                  Waypoint OP_PowderA_abov: TCP in base x=-12.145 y=-363.335 z=315.326 mm, rx=-0.7771 ry=1.753 rz=-1.7409 rad; joints [-58.232, -116.012, -83.989, -160.83, 75.01, 1.147] deg; TCP offset x=0 y=0 z=161 mm, rx=3.1415 ry=0 rz=0 rad
                  Waypoint OP_PowderA_pick: TCP in base x=-12.145 y=-363.335 z=179.899 mm, rx=-0.7771 ry=1.753 rz=-1.7409 rad; joints [-58.242, -124.732, -92.401, -143.702, 75.051, 1.161] deg
                  URCap Gripper (Robotiq_Grippers, Robotiq Inc.) dataModel(position=100.0, force=30.19607843137255, speed=30.19607843137255, positionInDouble=100.0, forceInDouble=30.19607843137255, speedInDouble=30.19607843137255, slaveIds=[9], blocking=true)
                  Wait Sleep waitTime=0.5
                  Set DigitalOutput pin=GRP_3F_Open; digitalValue=1
                  SuppressedNode
                    Script: Motors_off()
                  Waypoint OP_PowderA_abov: motionParameters(jointSpeed=1.047198 jointAcceleration=1.396263 cartesianSpeed=0.05 cartesianAcceleration=0.3); TCP in base x=-12.145 y=-363.335 z=315.326 mm, rx=-0.7771 ry=1.753 rz=-1.7409 rad; joints [-58.232, -116.012, -83.989, -160.83, 75.01, 1.147] deg
                  Waypoint Op_PowA_wP: TCP in base x=-173.728 y=-372.934 z=295.117 mm, rx=-0.9724 ry=1.541 rz=-1.5487 rad; joints [-67.269, -106.894, -99.849, -153.52, 49.211, 1.028] deg
              URCap Approach Pose (SensoPart VISOR Robotic, SensoPart Industriesensorik GmbH) dataModel(visorOffsetZ=0.0, visorJointSpeed=25.0, visorJointAcc=30.0); state(isChildrenLocked=true)
              URCap Target Pose (SensoPart VISOR Robotic, SensoPart Industriesensorik GmbH) dataModel(visorToolSpeed=50.0, visorToolAcc=100.0); state(isChildrenLocked=true)
              Folder Close Gripper
                target_pose := pose_add(get_actual_tcp_pose(), p[0,0,-0.1,0,0,0])
                MoveL speed 250 mm/s, acceleration 1200 mm/s^2 (useActiveTCP=true optimoveEnabled=false optiMoveSpeed=0.3 optiMoveAcceleration=0.09) feature=Base
                  Waypoint Variable (Variable): motionParameters(jointSpeed=1.047198 jointAcceleration=1.396263 cartesianSpeed=0.05 cartesianAcceleration=0.3); variable(name=target_pose)
                URCap Gripper (Robotiq_Grippers, Robotiq Inc.) dataModel(position=0.0, force=30.19607843137255, speed=30.19607843137255, positionInDouble=0.0, forceInDouble=30.19607843137255, speedInDouble=30.19607843137255, slaveIds=[9], blocking=true)
              URCap Exit Pose (SensoPart VISOR Robotic, SensoPart Industriesensorik GmbH) dataModel(visorOffsetZ=0.0); state(isChildrenLocked=true)
            URCap No Object Detected (SensoPart VISOR Robotic, SensoPart Industriesensorik GmbH) dataModel(Variable(key=visorNoObjCountVar, variable(name=easyPickNoObj_7, initializeExpression=0)))
              Popup Message (haltProgram=false message=No weigh scale detected inputType=Text)
        place_pose := get_actual_tcp_pose()
        Script: center_pose()
        SuppressedNode
          center_tilt_pos := P_center
        MoveJ speed 60 deg/s, acceleration 80 deg/s^2 (useActiveTCP=true optimoveEnabled=false optiMoveSpeed=0.3 optiMoveAcceleration=0.09) feature=Base
          Waypoint Waypoint_1: TCP in base x=-451.049 y=-340.589 z=308.224 mm, rx=0.0971 ry=0.091 rz=-1.5784 rad; joints [-127.334, -100.578, -80.109, -94.907, 86.186, -126.663] deg
    Case (caseValue=42)
      Folder Powder Emptying
        Script: zero_scale()
        Task := "Emptying"
        SuppressedNode
          URCap VISOR Robotic App (SensoPart VISOR Robotic, SensoPart Industriesensorik GmbH) dataModel(visorAppTemplate=1); state(isChildrenLocked=true)
            URCap Easy Pick Setup (SensoPart VISOR Robotic, SensoPart Industriesensorik GmbH) dataModel(visorId=0, visorSetJob=true, visorImageAcqSetup=2, visorCalibSetNo=9, visorDetector=1, visorOffsetSet=true, visorImageAcqSource=2, visorJobName=Weigh_target, visorSetupStatus=5, Pose(key=visorGripPose, Position(key=posePosition, Length(key=X value=-0.477246 unit=M), Length(key=Y value=0.05319 unit=M), Length(key=Z value=0.184004 unit=M)), Rotation(key=poseRotation, Angle(key=RX value=0.786642 unit=RAD), Angle(key=RY value=1.426517 unit=RAD), Angle(key=RZ value=-0.850311 unit=RAD))), Feature(key=visorImageAcqFeature name=FRM_Centrifuge)); state(isChildrenLocked=true)
            URCap Process (SensoPart VISOR Robotic, SensoPart Industriesensorik GmbH) dataModel(Variable(key=visorCounterVar, variable(name=easyPickCount_4, initializeExpression=0)), Variable(key=visorPartsFoundVar, variable(name=easyPickParts_4, initializeExpression=0))); state(isChildrenLocked=true)
              URCap Image Acquisition Pose (SensoPart VISOR Robotic, SensoPart Industriesensorik GmbH) state(isChildrenLocked=true)
              URCap Object Detected (SensoPart VISOR Robotic, SensoPart Industriesensorik GmbH) state(isChildrenLocked=true)
                Folder Open Gripper
                  Script: tare_scale()
                  Wait Sleep waitTime=0.2
                  Weight_value := get_weight()
                  Wait Sleep waitTime=0.2
                  Script: compute_level_percent(W_now, Weight_value)
                  If level≥10.0
                    MoveJ speed 60 deg/s, acceleration 80 deg/s^2 (useActiveTCP=true optimoveEnabled=false optiMoveSpeed=0.3 optiMoveAcceleration=0.09) feature=Base
                      Waypoint Spatula_otw: TCP in base x=-38.472 y=-263.141 z=425.351 mm, rx=-0.0004 ry=-0.0001 rz=3.0344 rad; joints [-68.119, -57.773, -97.702, -114.504, 90.127, 27.957] deg
                      Waypoint pick_spat_L_abv: TCP in base x=247.376 y=-151.301 z=298.406 mm, rx=0 ry=-0.0005 rz=3.0677 rad; joints [-4.058, -56.828, -117.366, -95.794, 90.156, 90.183] deg
                    MoveL speed 250 mm/s, acceleration 1200 mm/s^2 (useActiveTCP=true optimoveEnabled=false optiMoveSpeed=0.3 optiMoveAcceleration=0.09) feature=Base
                      Waypoint spat_L_pick: TCP in base x=244.425 y=-151.048 z=192.288 mm, rx=0 ry=-0.0005 rz=3.0677 rad; joints [-4.109, -56.947, -132.87, -80.171, 90.162, 90.196] deg
                      URCap Gripper (Robotiq_Grippers, Robotiq Inc.) dataModel(position=100.0, force=30.0, speed=0.0, positionInDouble=100.0, forceInDouble=30.0, speedInDouble=0.0, slaveIds=[9], blocking=true)
                      Waypoint spat_L_lift: TCP in base x=247.5 y=-151.291 z=242.147 mm, rx=0 ry=-0.0005 rz=3.0677 rad; joints [-4.086, -56.571, -125.696, -87.721, 90.161, 90.187] deg
                      Waypoint spat_L_side: TCP in base x=251.772 y=-93.61 z=242.166 mm, rx=0 ry=-0.0005 rz=3.0677 rad; joints [9.346, -52.481, -127.212, -90.293, 90.165, 103.617] deg
                      Waypoint spat_L_up: TCP in base x=248.632 y=-94.371 z=425.351 mm, rx=0 ry=-0.0005 rz=3.0677 rad; joints [9.417, -57.776, -97.699, -114.51, 90.125, 103.584] deg
                    MoveJ speed 60 deg/s, acceleration 80 deg/s^2 (useActiveTCP=true optimoveEnabled=false optiMoveSpeed=0.3 optiMoveAcceleration=0.09) feature=Base
                      Waypoint Spatula_otw: TCP in base x=-38.472 y=-263.141 z=425.351 mm, rx=-0.0004 ry=-0.0001 rz=3.0344 rad; joints [-68.119, -57.773, -97.702, -114.504, 90.127, 27.957] deg
                  ElseIf level≥1.0  and level<10.0
                    MoveJ speed 60 deg/s, acceleration 80 deg/s^2 (useActiveTCP=true optimoveEnabled=false optiMoveSpeed=0.3 optiMoveAcceleration=0.09) feature=Base
                      Waypoint Spatula_otw: TCP in base x=-38.472 y=-263.141 z=425.351 mm, rx=-0.0004 ry=-0.0001 rz=3.0344 rad; joints [-68.119, -57.773, -97.702, -114.504, 90.127, 27.957] deg
                      Waypoint spat_M_up: TCP in base x=246.651 y=-200.758 z=427.983 mm, rx=0 ry=-0.0005 rz=3.0677 rad; joints [-14.256, -65.249, -93.994, -110.748, 90.126, 79.91] deg
                    MoveL speed 250 mm/s, acceleration 1200 mm/s^2 (useActiveTCP=true optimoveEnabled=false optiMoveSpeed=0.3 optiMoveAcceleration=0.09) feature=Base
                      Waypoint spat_M_pick: TCP in base x=243.755 y=-195.91 z=192.274 mm, rx=0 ry=-0.0005 rz=3.0677 rad; joints [-13.585, -61.967, -130.669, -77.355, 90.156, 80.721] deg
                      URCap Gripper (Robotiq_Grippers, Robotiq Inc.) dataModel(position=100.0, force=30.0, speed=0.0, positionInDouble=100.0, forceInDouble=30.0, speedInDouble=0.0, slaveIds=[9], blocking=true)
                      Waypoint spat_M_up: TCP in base x=246.651 y=-200.758 z=427.983 mm, rx=0 ry=-0.0005 rz=3.0677 rad; joints [-14.256, -65.249, -93.994, -110.748, 90.126, 79.91] deg
                      Waypoint Spatula_otw: TCP in base x=-38.472 y=-263.141 z=425.351 mm, rx=-0.0004 ry=-0.0001 rz=3.0344 rad; joints [-68.119, -57.773, -97.702, -114.504, 90.127, 27.957] deg
                    switch_spat_M := False
                  Else 
                    MoveJ speed 60 deg/s, acceleration 80 deg/s^2 (useActiveTCP=true optimoveEnabled=false optiMoveSpeed=0.3 optiMoveAcceleration=0.09) feature=Base
                      Waypoint Spatula_otw: TCP in base x=-38.472 y=-263.141 z=425.351 mm, rx=-0.0004 ry=-0.0001 rz=3.0344 rad; joints [-68.119, -57.773, -97.702, -114.504, 90.127, 27.957] deg
                      Waypoint spat_S_up: TCP in base x=250.5 y=-246.906 z=391.584 mm, rx=0 ry=-0.0005 rz=3.0677 rad; joints [-22.233, -68.542, -97.739, -103.711, 90.135, 71.952] deg
                    MoveL speed 250 mm/s, acceleration 1200 mm/s^2 (useActiveTCP=true optimoveEnabled=false optiMoveSpeed=0.3 optiMoveAcceleration=0.09) feature=Base
                      Waypoint spat_S_pick: TCP in base x=245.173 y=-244.25 z=193.022 mm, rx=0 ry=-0.0005 rz=3.0677 rad; joints [-22.252, -68.068, -127.331, -74.593, 90.149, 72.053] deg
                      URCap Gripper (Robotiq_Grippers, Robotiq Inc.) dataModel(position=100.0, force=30.19607843137255, speed=0.0, positionInDouble=100.0, forceInDouble=30.19607843137255, speedInDouble=0.0, slaveIds=[9], blocking=true)
                      Waypoint spat_S_up: TCP in base x=250.5 y=-246.906 z=391.584 mm, rx=0 ry=-0.0005 rz=3.0677 rad; joints [-22.233, -68.542, -97.739, -103.711, 90.135, 71.952] deg
                      Waypoint Spatula_otw: TCP in base x=-38.472 y=-263.141 z=425.351 mm, rx=-0.0004 ry=-0.0001 rz=3.0344 rad; joints [-68.119, -57.773, -97.702, -114.504, 90.127, 27.957] deg
                    switch_spat_S := False
                  Weight_value := get_weight()
                  Script: auto_tilt_and_scoop(W_now, Target_weight, Weight_value)
                URCap Approach Pose (SensoPart VISOR Robotic, SensoPart Industriesensorik GmbH) dataModel(visorOffsetZ=-50.0, visorJointSpeed=10.0, visorJointAcc=15.0); state(isChildrenLocked=true)
                URCap Target Pose (SensoPart VISOR Robotic, SensoPart Industriesensorik GmbH) dataModel(visorToolSpeed=20.0, visorToolAcc=50.0); state(isChildrenLocked=true)
                Folder Close Gripper
                  dispense_pos := get_actual_tcp_pose()
                  Loop While (checkContinuously=false) expression=Weight_value≤Target_weight
                    MoveL speed 250 mm/s, acceleration 1200 mm/s^2 (useActiveTCP=true optimoveEnabled=false optiMoveSpeed=0.3 optiMoveAcceleration=0.09) feature=Base
                      Waypoint Variable (Variable): motionParameters(jointSpeed=0.436332 jointAcceleration=0.523599 cartesianSpeed=0.1 cartesianAcceleration=0.2); variable(name=dispense_pos)
                      Script: log_weight()
                      Wait Sleep waitTime=0.5
                      If level≥90.0
                        Script: Rotate()
                      If level≤70
                        Script: tilt_to_home()
                      Wait Sleep waitTime=0.5
                      Start_thread := True
                      vib_mot_thread := True
                      SuppressedNode
                        tilt_angle := current_pose[5]
                      Wait Sleep waitTime=0.5
                      SuppressedNode
                        Loop While (checkContinuously=true) expression=diff>3.0
                          tilt_pose := pose_trans(get_actual_tcp_pose(), p[0, 0, 0, 0, 0, 1.0])
                          Script: movel(tilt_pose, a=0.1, v=0.1, r=0.00001)
                          tilt_pose := pose_trans(get_actual_tcp_pose(), p[0, 0, 0, 0, 0, -1.0])
                          Script: movel(tilt_pose, a=0.1, v=0.1, r=0.00001)
                      If diff>0
                        tilt_pose := pose_trans(get_actual_tcp_pose(), p[0, 0, 0, 0, 0, 2.0])
                        Script: movel(tilt_pose, a=0.1, v=0.1, r=0.00001)
                      SuppressedNode
                        ElseIf diff≤1.0
                          Loop While (checkContinuously=false) expression=Weight_value≤Target_weight and tilt_angle≥(-1.999) and tilt_angle≤0.4
                            current_error := Target_weight-Weight_value
                            Integral_error := Integral_error+current_error*dt
                            derivative := (current_error-previous_error)/dt
                            tilt_increment := (kp*current_error)+(ki*Integral_error)+(kd*derivative)
                            current_pose := get_actual_tcp_pose()
                            tilt_angle := current_pose[5]
                            tilt_pose := pose_trans(current_pose, p[0, 0, 0, 0, 0, tilt_increment])
                            Script: movel(tilt_pose, a=0.1, v=0.1, r=0.00001)
                            previous_error := current_error
                      Start_thread := False
                      SuppressedNode
                        Waypoint Waypoint_64: motionParameters(jointSpeed=1.047198 jointAcceleration=1.396263 cartesianSpeed=0.03 cartesianAcceleration=0.1 blendRadius=0.05); TCP in base x=-542.998 y=-117.021 z=221.977 mm, rx=1.8981 ry=-0.7227 rz=1.5827 rad; joints [-123.845, -120.87, -101.018, -172.406, 14.907, 127.864] deg
                      Weight_value := get_weight()
                      SuppressedNode
                        tilt_angle := -1
                      Wait Sleep waitTime=0.5
                      vib_mot_thread := False
                      MoveL speed 250 mm/s, acceleration 500 mm/s^2 (useActiveTCP=true optimoveEnabled=false optiMoveSpeed=0.3 optiMoveAcceleration=0.09) feature=Base
                        Waypoint Variable (Variable): variable=dispense_pos
                      Integral_error := 0
                      current_error := 0
                      previous_error := 0
                      Set AnalogOutput pin=analog_out[0]; analogValue=0
                      Script: compute_level_percent(W_now, Weight_value)
                      If spatula ≟ "spatula_M"  and switch_spat_M≟ True
                        MoveJ speed 60 deg/s, acceleration 80 deg/s^2 (useActiveTCP=true optimoveEnabled=false optiMoveSpeed=0.3 optiMoveAcceleration=0.09) feature=Base
                          Waypoint Spatula_otw: TCP in base x=-38.472 y=-263.141 z=425.351 mm, rx=-0.0004 ry=-0.0001 rz=3.0344 rad; joints [-68.119, -57.773, -97.702, -114.504, 90.127, 27.957] deg
                          Waypoint spat_L_up: TCP in base x=248.632 y=-94.371 z=425.351 mm, rx=0 ry=-0.0005 rz=3.0677 rad; joints [9.417, -57.776, -97.699, -114.51, 90.125, 103.584] deg
                        MoveL speed 250 mm/s, acceleration 1200 mm/s^2 (useActiveTCP=true optimoveEnabled=false optiMoveSpeed=0.3 optiMoveAcceleration=0.09) feature=Base
                          Waypoint spat_L_side: TCP in base x=251.772 y=-93.61 z=242.166 mm, rx=0 ry=-0.0005 rz=3.0677 rad; joints [9.346, -52.481, -127.212, -90.293, 90.165, 103.617] deg
                          Waypoint spat_L_lift: TCP in base x=247.5 y=-151.291 z=242.147 mm, rx=0 ry=-0.0005 rz=3.0677 rad; joints [-4.086, -56.571, -125.696, -87.721, 90.161, 90.187] deg
                          Waypoint spat_L_pick: TCP in base x=244.425 y=-151.048 z=192.288 mm, rx=0 ry=-0.0005 rz=3.0677 rad; joints [-4.109, -56.947, -132.87, -80.171, 90.162, 90.196] deg
                          URCap Gripper (Robotiq_Grippers, Robotiq Inc.) dataModel(position=0.0, force=30.0, speed=100.0, positionInDouble=0.0, forceInDouble=30.0, speedInDouble=100.0, slaveIds=[9], blocking=true)
                          Waypoint spat_M_pick: TCP in base x=243.755 y=-195.91 z=192.274 mm, rx=0 ry=-0.0005 rz=3.0677 rad; joints [-13.585, -61.967, -130.669, -77.355, 90.156, 80.721] deg
                          URCap Gripper (Robotiq_Grippers, Robotiq Inc.) dataModel(position=100.0, force=30.0, speed=0.0, positionInDouble=100.0, forceInDouble=30.0, speedInDouble=0.0, slaveIds=[9], blocking=true)
                          Waypoint spat_M_up: TCP in base x=246.651 y=-200.758 z=427.983 mm, rx=0 ry=-0.0005 rz=3.0677 rad; joints [-14.256, -65.249, -93.994, -110.748, 90.126, 79.91] deg
                          Waypoint Spatula_otw: TCP in base x=-38.472 y=-263.141 z=425.351 mm, rx=-0.0004 ry=-0.0001 rz=3.0344 rad; joints [-68.119, -57.773, -97.702, -114.504, 90.127, 27.957] deg
                        switch_spat_M := False
                      ElseIf spatula ≟ "spatula_S" and switch_spat_S ≟ True
                        MoveL speed 250 mm/s, acceleration 1200 mm/s^2 (useActiveTCP=true optimoveEnabled=false optiMoveSpeed=0.3 optiMoveAcceleration=0.09) feature=Base
                          Waypoint Spatula_otw: TCP in base x=-38.472 y=-263.141 z=425.351 mm, rx=-0.0004 ry=-0.0001 rz=3.0344 rad; joints [-68.119, -57.773, -97.702, -114.504, 90.127, 27.957] deg
                          Waypoint spat_M_up: TCP in base x=246.651 y=-200.758 z=427.983 mm, rx=0 ry=-0.0005 rz=3.0677 rad; joints [-14.256, -65.249, -93.994, -110.748, 90.126, 79.91] deg
                          Waypoint spat_M_pick: TCP in base x=243.755 y=-195.91 z=192.274 mm, rx=0 ry=-0.0005 rz=3.0677 rad; joints [-13.585, -61.967, -130.669, -77.355, 90.156, 80.721] deg
                          URCap Gripper (Robotiq_Grippers, Robotiq Inc.) dataModel(position=0.0, force=30.19607843137255, speed=100.0, positionInDouble=0.0, forceInDouble=30.19607843137255, speedInDouble=100.0, slaveIds=[9], blocking=true)
                          Waypoint spat_S_pick: TCP in base x=245.173 y=-244.25 z=193.022 mm, rx=0 ry=-0.0005 rz=3.0677 rad; joints [-22.252, -68.068, -127.331, -74.593, 90.149, 72.053] deg
                          URCap Gripper (Robotiq_Grippers, Robotiq Inc.) dataModel(position=100.0, force=30.19607843137255, speed=0.0, positionInDouble=100.0, forceInDouble=30.19607843137255, speedInDouble=0.0, slaveIds=[9], blocking=true)
                          Waypoint spat_S_up: TCP in base x=250.5 y=-246.906 z=391.584 mm, rx=0 ry=-0.0005 rz=3.0677 rad; joints [-22.233, -68.542, -97.739, -103.711, 90.135, 71.952] deg
                          Waypoint Spatula_otw: TCP in base x=-38.472 y=-263.141 z=425.351 mm, rx=-0.0004 ry=-0.0001 rz=3.0344 rad; joints [-68.119, -57.773, -97.702, -114.504, 90.127, 27.957] deg
                        switch_spat_S := False
                      Script: auto_tilt_and_scoop(W_now, Target_weight, Weight_value)
                      Wait Sleep waitTime=0.5
                  SuppressedNode
                    Script: Rotate()
                URCap Exit Pose (SensoPart VISOR Robotic, SensoPart Industriesensorik GmbH) dataModel(visorOffsetZ=0.0); state(isChildrenLocked=true)
              URCap No Object Detected (SensoPart VISOR Robotic, SensoPart Industriesensorik GmbH) dataModel(Variable(key=visorNoObjCountVar, variable(name=easyPickNoObj_4, initializeExpression=0)))
                Popup Message (haltProgram=false message=No weigh scale detected inputType=Text)
        SuppressedNode
          Folder powder dispensing
            SuppressedNode
              Target_weight := Target_weight/1000
            Loop While (checkContinuously=false) expression=Weight_value<Target_weight
              Script: auto_tilt_and_scoop(W_now, Target_weight, Weight_value)
              Start_thread := True
              MoveL speed 250 mm/s, acceleration 1200 mm/s^2 (useActiveTCP=true optimoveEnabled=false optiMoveSpeed=0.3 optiMoveAcceleration=0.09) feature=Base
                Waypoint Variable (Variable): motionParameters(jointSpeed=0.436332 jointAcceleration=0.523599 cartesianSpeed=0.05 cartesianAcceleration=0.2); variable=dispense_pos
                Wait Sleep waitTime=0.5
                Script: Rotate()
                Wait Sleep waitTime=0.5
              MoveL speed 250 mm/s, acceleration 1200 mm/s^2 (useActiveTCP=true optimoveEnabled=false optiMoveSpeed=0.3 optiMoveAcceleration=0.09) feature=Base
                Start_thread := True
                vib_mot_thread := True
                tilt_angle := current_pose[5]
                Wait Sleep waitTime=0.5
                SuppressedNode
                  Loop While (checkContinuously=true) expression=diff>3.0
                    tilt_pose := pose_trans(get_actual_tcp_pose(), p[0, 0, 0, 0, 0, 1.0])
                    Script: movel(tilt_pose, a=0.1, v=0.1, r=0.00001)
                    tilt_pose := pose_trans(get_actual_tcp_pose(), p[0, 0, 0, 0, 0, -1.0])
                    Script: movel(tilt_pose, a=0.1, v=0.1, r=0.00001)
                If diff>3.0
                  tilt_pose := pose_trans(get_actual_tcp_pose(), p[0, 0, 0, 0, 0, 2.0])
                  Script: movel(tilt_pose, a=0.1, v=0.1, r=0.00001)
                ElseIf diff≤3.0
                  Loop While (checkContinuously=false) expression=Weight_value≤Target_weight and tilt_angle≥(-1.999) and tilt_angle≤0
                    current_error := Target_weight-Weight_value
                    Integral_error := Integral_error+current_error*dt
                    derivative := (current_error-previous_error)/dt
                    tilt_increment := (kp*current_error)+(ki*Integral_error)+(kd*derivative)
                    current_pose := get_actual_tcp_pose()
                    tilt_angle := current_pose[5]
                    tilt_pose := pose_trans(current_pose, p[0, 0, 0, 0, 0, tilt_increment])
                    Script: movel(tilt_pose, a=0.1, v=0.1, r=0.00001)
                    previous_error := current_error
                Start_thread := False
                SuppressedNode
                  Waypoint Waypoint_64: motionParameters(jointSpeed=1.047198 jointAcceleration=1.396263 cartesianSpeed=0.03 cartesianAcceleration=0.1 blendRadius=0.05); TCP in base x=-542.998 y=-117.021 z=221.977 mm, rx=1.8981 ry=-0.7227 rz=1.5827 rad; joints [-123.845, -120.87, -101.018, -172.406, 14.907, 127.864] deg
                Weight_value := get_weight()
                Wait Sleep waitTime=0.5
                tilt_angle := -1
                vib_mot_thread := False
                MoveL speed 50 mm/s, acceleration 300 mm/s^2 (useActiveTCP=true optimoveEnabled=false optiMoveSpeed=0.3 optiMoveAcceleration=0.09) feature=Base
                  Waypoint Variable (Variable): motionParameters(jointSpeed=0.436332 jointAcceleration=0.523599 cartesianSpeed=0.05 cartesianAcceleration=0.2); variable=dispense_pos
                Integral_error := 0
                current_error := 0
                previous_error := 0
                Set AnalogOutput pin=analog_out[0]; analogValue=0
              Script: movel(pose_trans(dispense_pos, p[-0.02,0,0,0,0,0]))
            SuppressedNode
              MoveL speed 250 mm/s, acceleration 1200 mm/s^2 (useActiveTCP=true optimoveEnabled=false optiMoveSpeed=0.3 optiMoveAcceleration=0.09) feature=Base
                Waypoint aftr_scoo3: motionParameters(jointSpeed=1.047198 jointAcceleration=1.396263 cartesianSpeed=0.1 cartesianAcceleration=0.3); TCP in base x=-289.76 y=-315.385 z=303.744 mm, rx=0.16 ry=1.6274 rz=-0.3449 rad; joints [-76.632, -96.313, -113.776, -155.476, 32.027, -78.1] deg
                Waypoint ftr_scoop2: motionParameters(jointSpeed=1.047198 jointAcceleration=1.396263 cartesianSpeed=0.1 cartesianAcceleration=0.4); TCP in base x=194.287 y=-495.78 z=282.072 mm, rx=-0.179 ry=1.6121 rz=-0.016 rad; joints [-34.133, -129.723, -68.393, -165.549, 50.138, -80.843] deg
                Waypoint aftr_scoop1: motionParameters(jointSpeed=1.047198 jointAcceleration=1.396263 cartesianSpeed=0.1 cartesianAcceleration=0.4); TCP in base x=138.504 y=-514.48 z=214.154 mm, rx=-0.1348 ry=1.5599 rz=-0.0592 rad; joints [-39.422, -130.004, -76.262, -153.157, 47.788, -83.41] deg
                Waypoint After_disp_3: motionParameters(jointSpeed=1.047198 jointAcceleration=1.396263 cartesianSpeed=0.1 cartesianAcceleration=0.4); TCP in base x=125.935 y=-585.611 z=299.546 mm, rx=0.9596 ry=-0.1344 rz=2.8807 rad; joints [-54.056, -115.535, -63.235, -120.118, 65.773, 48.319] deg
                Set AnalogOutput pin=analog_out[0]; analogValue=3
                Wait Sleep waitTime=2
                Set AnalogOutput pin=analog_out[0]; analogValue=0
                Waypoint aftr_scoop1: TCP in base x=138.504 y=-514.48 z=214.154 mm, rx=-0.1348 ry=1.5599 rz=-0.0592 rad; joints [-39.422, -130.004, -76.262, -153.157, 47.788, -83.41] deg
                Waypoint ftr_scoop2: motionParameters(jointSpeed=1.047198 jointAcceleration=1.396263 cartesianSpeed=0.1 cartesianAcceleration=0.4); TCP in base x=194.287 y=-495.78 z=282.072 mm, rx=-0.179 ry=1.6121 rz=-0.016 rad; joints [-34.133, -129.723, -68.393, -165.549, 50.138, -80.843] deg
                Waypoint Waypoint_63: motionParameters(blendRadius=0.05); TCP in base x=101.295 y=-465.376 z=381.756 mm, rx=0.9726 ry=-0.1584 rz=2.8872 rad; joints [-48.863, -99.659, -71.872, -130.079, 68.56, 52.636] deg; TCP offset x=0 y=0 z=161 mm, rx=3.1415 ry=0 rz=0 rad
                Waypoint Start: motionParameters(jointSpeed=1.047198 jointAcceleration=1.396263 cartesianSpeed=0.15 cartesianAcceleration=0.6); TCP in base x=-33.065 y=-365.399 z=389.873 mm, rx=0 ry=0 rz=2.7258 rad; joints [-73.774, -70.638, -96.716, -102.629, 90.121, 40.001] deg; TCP offset x=0 y=0 z=161 mm, rx=3.1415 ry=0 rz=0 rad
                Popup Message (haltProgram=false message=Powder dispensed successfully... inputType=Text)
            SuppressedNode
              Script: tilt()
        SuppressedNode
          Script: tilt_send()
    Case (caseValue=43)
      Folder Powder dosing
        Script: zero_scale()
        SuppressedNode
          URCap VISOR Robotic App (SensoPart VISOR Robotic, SensoPart Industriesensorik GmbH) dataModel(visorAppTemplate=1); state(isChildrenLocked=true)
            URCap Easy Pick Setup (SensoPart VISOR Robotic, SensoPart Industriesensorik GmbH) dataModel(visorId=0, visorSetJob=true, visorImageAcqSetup=2, visorCalibSetNo=9, visorDetector=1, visorOffsetSet=true, visorImageAcqSource=2, visorJobName=Weigh_target, visorSetupStatus=5, Pose(key=visorGripPose, Position(key=posePosition, Length(key=X value=-0.477246 unit=M), Length(key=Y value=0.05319 unit=M), Length(key=Z value=0.184004 unit=M)), Rotation(key=poseRotation, Angle(key=RX value=0.786642 unit=RAD), Angle(key=RY value=1.426517 unit=RAD), Angle(key=RZ value=-0.850311 unit=RAD))), Feature(key=visorImageAcqFeature name=FRM_Centrifuge)); state(isChildrenLocked=true)
            URCap Process (SensoPart VISOR Robotic, SensoPart Industriesensorik GmbH) dataModel(Variable(key=visorCounterVar, variable(name=easyPickCount_4, initializeExpression=0)), Variable(key=visorPartsFoundVar, variable(name=easyPickParts_4, initializeExpression=0))); state(isChildrenLocked=true)
              URCap Image Acquisition Pose (SensoPart VISOR Robotic, SensoPart Industriesensorik GmbH) state(isChildrenLocked=true)
              URCap Object Detected (SensoPart VISOR Robotic, SensoPart Industriesensorik GmbH) state(isChildrenLocked=true)
                Folder Open Gripper
                  Script: tare_scale()
                  Wait Sleep waitTime=0.2
                  Weight_value := get_weight()
                  Wait Sleep waitTime=0.2
                  diff := Target_weight-Weight_value
                  Script: compute_level_percent(W_now, Weight_value)
                  Script: spatula = select_spatula(Pow_name, level, diff)
                  If spatula ≟ "spatula_L"
                    MoveJ speed 60 deg/s, acceleration 80 deg/s^2 (useActiveTCP=true optimoveEnabled=false optiMoveSpeed=0.3 optiMoveAcceleration=0.09) feature=Base
                      Waypoint Spatula_otw: TCP in base x=-38.472 y=-263.141 z=425.351 mm, rx=-0.0004 ry=-0.0001 rz=3.0344 rad; joints [-68.119, -57.773, -97.702, -114.504, 90.127, 27.957] deg
                      Waypoint pick_spat_L_abv: TCP in base x=247.376 y=-151.301 z=298.406 mm, rx=0 ry=-0.0005 rz=3.0677 rad; joints [-4.058, -56.828, -117.366, -95.794, 90.156, 90.183] deg
                    MoveL speed 250 mm/s, acceleration 1200 mm/s^2 (useActiveTCP=true optimoveEnabled=false optiMoveSpeed=0.3 optiMoveAcceleration=0.09) feature=Base
                      Waypoint spat_L_pick: TCP in base x=244.425 y=-151.048 z=192.288 mm, rx=0 ry=-0.0005 rz=3.0677 rad; joints [-4.109, -56.947, -132.87, -80.171, 90.162, 90.196] deg
                      URCap Gripper (Robotiq_Grippers, Robotiq Inc.) dataModel(position=100.0, force=30.0, speed=0.0, positionInDouble=100.0, forceInDouble=30.0, speedInDouble=0.0, slaveIds=[9], blocking=true)
                      Waypoint spat_L_lift: TCP in base x=247.5 y=-151.291 z=242.147 mm, rx=0 ry=-0.0005 rz=3.0677 rad; joints [-4.086, -56.571, -125.696, -87.721, 90.161, 90.187] deg
                      Waypoint spat_L_side: TCP in base x=251.772 y=-93.61 z=242.166 mm, rx=0 ry=-0.0005 rz=3.0677 rad; joints [9.346, -52.481, -127.212, -90.293, 90.165, 103.617] deg
                      Waypoint spat_L_up: TCP in base x=248.632 y=-94.371 z=425.351 mm, rx=0 ry=-0.0005 rz=3.0677 rad; joints [9.417, -57.776, -97.699, -114.51, 90.125, 103.584] deg
                    MoveJ speed 60 deg/s, acceleration 80 deg/s^2 (useActiveTCP=true optimoveEnabled=false optiMoveSpeed=0.3 optiMoveAcceleration=0.09) feature=Base
                      Waypoint Spatula_otw: TCP in base x=-38.472 y=-263.141 z=425.351 mm, rx=-0.0004 ry=-0.0001 rz=3.0344 rad; joints [-68.119, -57.773, -97.702, -114.504, 90.127, 27.957] deg
                  ElseIf spatula ≟"spatula_M"
                    MoveJ speed 60 deg/s, acceleration 80 deg/s^2 (useActiveTCP=true optimoveEnabled=false optiMoveSpeed=0.3 optiMoveAcceleration=0.09) feature=Base
                      Waypoint Spatula_otw: TCP in base x=-38.472 y=-263.141 z=425.351 mm, rx=-0.0004 ry=-0.0001 rz=3.0344 rad; joints [-68.119, -57.773, -97.702, -114.504, 90.127, 27.957] deg
                      Waypoint spat_M_up: TCP in base x=246.651 y=-200.758 z=427.983 mm, rx=0 ry=-0.0005 rz=3.0677 rad; joints [-14.256, -65.249, -93.994, -110.748, 90.126, 79.91] deg
                    MoveL speed 250 mm/s, acceleration 1200 mm/s^2 (useActiveTCP=true optimoveEnabled=false optiMoveSpeed=0.3 optiMoveAcceleration=0.09) feature=Base
                      Waypoint spat_M_pick: TCP in base x=243.755 y=-195.91 z=192.274 mm, rx=0 ry=-0.0005 rz=3.0677 rad; joints [-13.585, -61.967, -130.669, -77.355, 90.156, 80.721] deg
                      URCap Gripper (Robotiq_Grippers, Robotiq Inc.) dataModel(position=100.0, force=30.0, speed=0.0, positionInDouble=100.0, forceInDouble=30.0, speedInDouble=0.0, slaveIds=[9], blocking=true)
                      Waypoint spat_M_up: TCP in base x=246.651 y=-200.758 z=427.983 mm, rx=0 ry=-0.0005 rz=3.0677 rad; joints [-14.256, -65.249, -93.994, -110.748, 90.126, 79.91] deg
                      Waypoint Spatula_otw: TCP in base x=-38.472 y=-263.141 z=425.351 mm, rx=-0.0004 ry=-0.0001 rz=3.0344 rad; joints [-68.119, -57.773, -97.702, -114.504, 90.127, 27.957] deg
                    switch_spat_M := False
                  ElseIf spatula≟"spatula_S"
                    MoveJ speed 60 deg/s, acceleration 80 deg/s^2 (useActiveTCP=true optimoveEnabled=false optiMoveSpeed=0.3 optiMoveAcceleration=0.09) feature=Base
                      Waypoint Spatula_otw: TCP in base x=-38.472 y=-263.141 z=425.351 mm, rx=-0.0004 ry=-0.0001 rz=3.0344 rad; joints [-68.119, -57.773, -97.702, -114.504, 90.127, 27.957] deg
                      Waypoint spat_M_up: TCP in base x=246.651 y=-200.758 z=427.983 mm, rx=0 ry=-0.0005 rz=3.0677 rad; joints [-14.256, -65.249, -93.994, -110.748, 90.126, 79.91] deg
                    MoveL speed 250 mm/s, acceleration 1200 mm/s^2 (useActiveTCP=true optimoveEnabled=false optiMoveSpeed=0.3 optiMoveAcceleration=0.09) feature=Base
                      Waypoint spat_M_pick: TCP in base x=243.755 y=-195.91 z=192.274 mm, rx=0 ry=-0.0005 rz=3.0677 rad; joints [-13.585, -61.967, -130.669, -77.355, 90.156, 80.721] deg
                      URCap Gripper (Robotiq_Grippers, Robotiq Inc.) dataModel(position=100.0, force=30.0, speed=0.0, positionInDouble=100.0, forceInDouble=30.0, speedInDouble=0.0, slaveIds=[9], blocking=true)
                      Waypoint spat_M_up: TCP in base x=246.651 y=-200.758 z=427.983 mm, rx=0 ry=-0.0005 rz=3.0677 rad; joints [-14.256, -65.249, -93.994, -110.748, 90.126, 79.91] deg
                      Waypoint Spatula_otw: TCP in base x=-38.472 y=-263.141 z=425.351 mm, rx=-0.0004 ry=-0.0001 rz=3.0344 rad; joints [-68.119, -57.773, -97.702, -114.504, 90.127, 27.957] deg
                    switch_spat_M := False
                  Weight_value := get_weight()
                  Script: auto_tilt_and_scoop(W_now, Target_weight, Weight_value)
                URCap Approach Pose (SensoPart VISOR Robotic, SensoPart Industriesensorik GmbH) dataModel(visorOffsetZ=-50.0, visorJointSpeed=10.0, visorJointAcc=15.0); state(isChildrenLocked=true)
                URCap Target Pose (SensoPart VISOR Robotic, SensoPart Industriesensorik GmbH) dataModel(visorToolSpeed=20.0, visorToolAcc=50.0); state(isChildrenLocked=true)
                Folder Close Gripper
                  dispense_pos := get_actual_tcp_pose()
                  Loop While (checkContinuously=true) expression=Weight_value≤Target_weight
                    MoveL speed 250 mm/s, acceleration 1200 mm/s^2 (useActiveTCP=true optimoveEnabled=false optiMoveSpeed=0.3 optiMoveAcceleration=0.09) feature=Base
                      Waypoint Variable (Variable): motionParameters(jointSpeed=0.436332 jointAcceleration=0.523599 cartesianSpeed=0.1 cartesianAcceleration=0.2); variable=dispense_pos
                      Script: log_weight()
                      Wait Sleep waitTime=0.5
                      If level≥90.0
                        Script: Rotate()
                      If level≤70
                        Script: tilt_to_home()
                      Wait Sleep waitTime=0.5
                      Start_thread := True
                      vib_mot_thread := True
                      SuppressedNode
                        tilt_angle := current_pose[5]
                      Wait Sleep waitTime=0.5
                      SuppressedNode
                        Loop While (checkContinuously=true) expression=diff>3.0
                          tilt_pose := pose_trans(get_actual_tcp_pose(), p[0, 0, 0, 0, 0, 1.0])
                          Script: movel(tilt_pose, a=0.1, v=0.1, r=0.00001)
                          tilt_pose := pose_trans(get_actual_tcp_pose(), p[0, 0, 0, 0, 0, -1.0])
                          Script: movel(tilt_pose, a=0.1, v=0.1, r=0.00001)
                      If spatula ≟ "spatula_L"  and diff ≥3.5
                        tilt_pose := pose_trans(get_actual_tcp_pose(), p[0, 0, 0, 0, 0, 2.0])
                        Script: movel(tilt_pose, a=0.1, v=0.1, r=0.00001)
                      SuppressedNode
                        ElseIf diff≤1.0
                          Loop While (checkContinuously=false) expression=Weight_value≤Target_weight and tilt_angle≥(-1.999) and tilt_angle≤0.4
                            current_error := Target_weight-Weight_value
                            Integral_error := Integral_error+current_error*dt
                            derivative := (current_error-previous_error)/dt
                            tilt_increment := (kp*current_error)+(ki*Integral_error)+(kd*derivative)
                            current_pose := get_actual_tcp_pose()
                            tilt_angle := current_pose[5]
                            tilt_pose := pose_trans(current_pose, p[0, 0, 0, 0, 0, tilt_increment])
                            Script: movel(tilt_pose, a=0.1, v=0.1, r=0.00001)
                            previous_error := current_error
                      If spatula ≟ "spatula_M"  and diff ≥1.0
                        tilt_pose := pose_trans(get_actual_tcp_pose(), p[0, 0, 0, 0, 0, 2.0])
                        Script: movel(tilt_pose, a=0.1, v=0.1, r=0.00001)
                      ElseIf diff≤1.0
                        Loop While (checkContinuously=false) expression=Weight_value≤Target_weight and tilt_angle≥(-1.999) and tilt_angle≤0.5
                          current_error := Target_weight-Weight_value
                          Integral_error := Integral_error+current_error*dt
                          derivative := (current_error-previous_error)/dt
                          tilt_increment := (kp*current_error)+(ki*Integral_error)+(kd*derivative)
                          current_pose := get_actual_tcp_pose()
                          tilt_angle := current_pose[5]
                          tilt_pose := pose_trans(current_pose, p[0, 0, 0, 0, 0, tilt_increment])
                          Script: movel(tilt_pose, a=0.1, v=0.1, r=0.00001)
                          previous_error := current_error
                      Start_thread := False
                      SuppressedNode
                        Waypoint Waypoint_64: motionParameters(jointSpeed=1.047198 jointAcceleration=1.396263 cartesianSpeed=0.03 cartesianAcceleration=0.1 blendRadius=0.05); TCP in base x=-542.998 y=-117.021 z=221.977 mm, rx=1.8981 ry=-0.7227 rz=1.5827 rad; joints [-123.845, -120.87, -101.018, -172.406, 14.907, 127.864] deg
                      Weight_value := get_weight()
                      SuppressedNode
                        tilt_angle := -1
                      Wait Sleep waitTime=0.5
                      vib_mot_thread := False
                      MoveL speed 250 mm/s, acceleration 500 mm/s^2 (useActiveTCP=true optimoveEnabled=false optiMoveSpeed=0.3 optiMoveAcceleration=0.09) feature=Base
                        Waypoint Variable (Variable): variable=dispense_pos
                      Integral_error := 0
                      current_error := 0
                      previous_error := 0
                      Set AnalogOutput pin=analog_out[0]; analogValue=0
                      Script: select_spatula(Pow_name, level, diff)
                      If spatula ≟ "spatula_M"  and switch_spat_M≟ True
                        MoveJ speed 60 deg/s, acceleration 80 deg/s^2 (useActiveTCP=true optimoveEnabled=false optiMoveSpeed=0.3 optiMoveAcceleration=0.09) feature=Base
                          Waypoint Spatula_otw: TCP in base x=-38.472 y=-263.141 z=425.351 mm, rx=-0.0004 ry=-0.0001 rz=3.0344 rad; joints [-68.119, -57.773, -97.702, -114.504, 90.127, 27.957] deg
                          Waypoint spat_L_up: TCP in base x=248.632 y=-94.371 z=425.351 mm, rx=0 ry=-0.0005 rz=3.0677 rad; joints [9.417, -57.776, -97.699, -114.51, 90.125, 103.584] deg
                        MoveL speed 250 mm/s, acceleration 1200 mm/s^2 (useActiveTCP=true optimoveEnabled=false optiMoveSpeed=0.3 optiMoveAcceleration=0.09) feature=Base
                          Waypoint spat_L_side: TCP in base x=251.772 y=-93.61 z=242.166 mm, rx=0 ry=-0.0005 rz=3.0677 rad; joints [9.346, -52.481, -127.212, -90.293, 90.165, 103.617] deg
                          Waypoint spat_L_lift: TCP in base x=247.5 y=-151.291 z=242.147 mm, rx=0 ry=-0.0005 rz=3.0677 rad; joints [-4.086, -56.571, -125.696, -87.721, 90.161, 90.187] deg
                          Waypoint spat_L_pick: TCP in base x=244.425 y=-151.048 z=192.288 mm, rx=0 ry=-0.0005 rz=3.0677 rad; joints [-4.109, -56.947, -132.87, -80.171, 90.162, 90.196] deg
                          URCap Gripper (Robotiq_Grippers, Robotiq Inc.) dataModel(position=0.0, force=30.0, speed=100.0, positionInDouble=0.0, forceInDouble=30.0, speedInDouble=100.0, slaveIds=[9], blocking=true)
                          Waypoint spat_M_pick: TCP in base x=243.755 y=-195.91 z=192.274 mm, rx=0 ry=-0.0005 rz=3.0677 rad; joints [-13.585, -61.967, -130.669, -77.355, 90.156, 80.721] deg
                          URCap Gripper (Robotiq_Grippers, Robotiq Inc.) dataModel(position=100.0, force=30.0, speed=0.0, positionInDouble=100.0, forceInDouble=30.0, speedInDouble=0.0, slaveIds=[9], blocking=true)
                          Waypoint spat_M_up: TCP in base x=246.651 y=-200.758 z=427.983 mm, rx=0 ry=-0.0005 rz=3.0677 rad; joints [-14.256, -65.249, -93.994, -110.748, 90.126, 79.91] deg
                          Waypoint Spatula_otw: TCP in base x=-38.472 y=-263.141 z=425.351 mm, rx=-0.0004 ry=-0.0001 rz=3.0344 rad; joints [-68.119, -57.773, -97.702, -114.504, 90.127, 27.957] deg
                        switch_spat_M := False
                      ElseIf spatula ≟ "spatula_S" and switch_spat_S ≟ True
                        MoveL speed 250 mm/s, acceleration 1200 mm/s^2 (useActiveTCP=true optimoveEnabled=false optiMoveSpeed=0.3 optiMoveAcceleration=0.09) feature=Base
                          Waypoint Spatula_otw: TCP in base x=-38.472 y=-263.141 z=425.351 mm, rx=-0.0004 ry=-0.0001 rz=3.0344 rad; joints [-68.119, -57.773, -97.702, -114.504, 90.127, 27.957] deg
                          Waypoint spat_M_up: TCP in base x=246.651 y=-200.758 z=427.983 mm, rx=0 ry=-0.0005 rz=3.0677 rad; joints [-14.256, -65.249, -93.994, -110.748, 90.126, 79.91] deg
                          Waypoint spat_M_pick: TCP in base x=243.755 y=-195.91 z=192.274 mm, rx=0 ry=-0.0005 rz=3.0677 rad; joints [-13.585, -61.967, -130.669, -77.355, 90.156, 80.721] deg
                          URCap Gripper (Robotiq_Grippers, Robotiq Inc.) dataModel(position=0.0, force=30.19607843137255, speed=100.0, positionInDouble=0.0, forceInDouble=30.19607843137255, speedInDouble=100.0, slaveIds=[9], blocking=true)
                          Waypoint spat_S_pick: TCP in base x=245.173 y=-244.25 z=193.022 mm, rx=0 ry=-0.0005 rz=3.0677 rad; joints [-22.252, -68.068, -127.331, -74.593, 90.149, 72.053] deg
                          URCap Gripper (Robotiq_Grippers, Robotiq Inc.) dataModel(position=100.0, force=30.19607843137255, speed=0.0, positionInDouble=100.0, forceInDouble=30.19607843137255, speedInDouble=0.0, slaveIds=[9], blocking=true)
                          Waypoint spat_S_up: TCP in base x=250.5 y=-246.906 z=391.584 mm, rx=0 ry=-0.0005 rz=3.0677 rad; joints [-22.233, -68.542, -97.739, -103.711, 90.135, 71.952] deg
                          Waypoint Spatula_otw: TCP in base x=-38.472 y=-263.141 z=425.351 mm, rx=-0.0004 ry=-0.0001 rz=3.0344 rad; joints [-68.119, -57.773, -97.702, -114.504, 90.127, 27.957] deg
                        switch_spat_S := False
                      Script: auto_tilt_and_scoop(W_now, Target_weight, Weight_value)
                      Wait Sleep waitTime=0.5
                  Start_thread := False
                  Wait Sleep waitTime=0.5
                  vib_mot_thread := False
                  SuppressedNode
                    Script: Rotate()
                URCap Exit Pose (SensoPart VISOR Robotic, SensoPart Industriesensorik GmbH) dataModel(visorOffsetZ=0.0); state(isChildrenLocked=true)
              URCap No Object Detected (SensoPart VISOR Robotic, SensoPart Industriesensorik GmbH) dataModel(Variable(key=visorNoObjCountVar, variable(name=easyPickNoObj_4, initializeExpression=0)))
                Popup Message (haltProgram=false message=No weigh scale detected inputType=Text)
        Task := "Dosing"
        Script: scooping_init()
        SuppressedNode
          MoveJ speed 60 deg/s, acceleration 80 deg/s^2 (useActiveTCP=true optimoveEnabled=false optiMoveSpeed=0.3 optiMoveAcceleration=0.09) feature=Base
            Waypoint Variable (Variable): motionParameters(jointSpeed=0.436332 jointAcceleration=0.523599 cartesianSpeed=0.1 cartesianAcceleration=0.2); variable=dispense_pos
        Script: after_scoop()
        SuppressedNode
          Folder powder dispensing
            SuppressedNode
              Target_weight := Target_weight/1000
            Loop While (checkContinuously=false) expression=Weight_value<Target_weight
              Script: auto_tilt_and_scoop(W_now, Target_weight, Weight_value)
              Start_thread := True
              MoveL speed 250 mm/s, acceleration 1200 mm/s^2 (useActiveTCP=true optimoveEnabled=false optiMoveSpeed=0.3 optiMoveAcceleration=0.09) feature=Base
                Waypoint Variable (Variable): motionParameters(jointSpeed=0.436332 jointAcceleration=0.523599 cartesianSpeed=0.05 cartesianAcceleration=0.2); variable=dispense_pos
                Wait Sleep waitTime=0.5
                Script: Rotate()
                Wait Sleep waitTime=0.5
              MoveL speed 250 mm/s, acceleration 1200 mm/s^2 (useActiveTCP=true optimoveEnabled=false optiMoveSpeed=0.3 optiMoveAcceleration=0.09) feature=Base
                Start_thread := True
                vib_mot_thread := True
                tilt_angle := current_pose[5]
                Wait Sleep waitTime=0.5
                SuppressedNode
                  Loop While (checkContinuously=true) expression=diff>3.0
                    tilt_pose := pose_trans(get_actual_tcp_pose(), p[0, 0, 0, 0, 0, 1.0])
                    Script: movel(tilt_pose, a=0.1, v=0.1, r=0.00001)
                    tilt_pose := pose_trans(get_actual_tcp_pose(), p[0, 0, 0, 0, 0, -1.0])
                    Script: movel(tilt_pose, a=0.1, v=0.1, r=0.00001)
                If diff>3.0
                  tilt_pose := pose_trans(get_actual_tcp_pose(), p[0, 0, 0, 0, 0, 2.0])
                  Script: movel(tilt_pose, a=0.1, v=0.1, r=0.00001)
                ElseIf diff≤3.0
                  Loop While (checkContinuously=false) expression=Weight_value≤Target_weight and tilt_angle≥(-1.999) and tilt_angle≤0
                    current_error := Target_weight-Weight_value
                    Integral_error := Integral_error+current_error*dt
                    derivative := (current_error-previous_error)/dt
                    tilt_increment := (kp*current_error)+(ki*Integral_error)+(kd*derivative)
                    current_pose := get_actual_tcp_pose()
                    tilt_angle := current_pose[5]
                    tilt_pose := pose_trans(current_pose, p[0, 0, 0, 0, 0, tilt_increment])
                    Script: movel(tilt_pose, a=0.1, v=0.1, r=0.00001)
                    previous_error := current_error
                Start_thread := False
                SuppressedNode
                  Waypoint Waypoint_64: motionParameters(jointSpeed=1.047198 jointAcceleration=1.396263 cartesianSpeed=0.03 cartesianAcceleration=0.1 blendRadius=0.05); TCP in base x=-542.998 y=-117.021 z=221.977 mm, rx=1.8981 ry=-0.7227 rz=1.5827 rad; joints [-123.845, -120.87, -101.018, -172.406, 14.907, 127.864] deg
                Weight_value := get_weight()
                Wait Sleep waitTime=0.5
                tilt_angle := -1
                vib_mot_thread := False
                MoveL speed 50 mm/s, acceleration 300 mm/s^2 (useActiveTCP=true optimoveEnabled=false optiMoveSpeed=0.3 optiMoveAcceleration=0.09) feature=Base
                  Waypoint Variable (Variable): motionParameters(jointSpeed=0.436332 jointAcceleration=0.523599 cartesianSpeed=0.05 cartesianAcceleration=0.2); variable=dispense_pos
                Integral_error := 0
                current_error := 0
                previous_error := 0
                Set AnalogOutput pin=analog_out[0]; analogValue=0
              Script: movel(pose_trans(dispense_pos, p[-0.02,0,0,0,0,0]))
            SuppressedNode
              MoveL speed 250 mm/s, acceleration 1200 mm/s^2 (useActiveTCP=true optimoveEnabled=false optiMoveSpeed=0.3 optiMoveAcceleration=0.09) feature=Base
                Waypoint aftr_scoo3: motionParameters(jointSpeed=1.047198 jointAcceleration=1.396263 cartesianSpeed=0.1 cartesianAcceleration=0.3); TCP in base x=-289.76 y=-315.385 z=303.744 mm, rx=0.16 ry=1.6274 rz=-0.3449 rad; joints [-76.632, -96.313, -113.776, -155.476, 32.027, -78.1] deg
                Waypoint ftr_scoop2: motionParameters(jointSpeed=1.047198 jointAcceleration=1.396263 cartesianSpeed=0.1 cartesianAcceleration=0.4); TCP in base x=194.287 y=-495.78 z=282.072 mm, rx=-0.179 ry=1.6121 rz=-0.016 rad; joints [-34.133, -129.723, -68.393, -165.549, 50.138, -80.843] deg
                Waypoint aftr_scoop1: motionParameters(jointSpeed=1.047198 jointAcceleration=1.396263 cartesianSpeed=0.1 cartesianAcceleration=0.4); TCP in base x=138.504 y=-514.48 z=214.154 mm, rx=-0.1348 ry=1.5599 rz=-0.0592 rad; joints [-39.422, -130.004, -76.262, -153.157, 47.788, -83.41] deg
                Waypoint After_disp_3: motionParameters(jointSpeed=1.047198 jointAcceleration=1.396263 cartesianSpeed=0.1 cartesianAcceleration=0.4); TCP in base x=125.935 y=-585.611 z=299.546 mm, rx=0.9596 ry=-0.1344 rz=2.8807 rad; joints [-54.056, -115.535, -63.235, -120.118, 65.773, 48.319] deg
                Set AnalogOutput pin=analog_out[0]; analogValue=3
                Wait Sleep waitTime=2
                Set AnalogOutput pin=analog_out[0]; analogValue=0
                Waypoint aftr_scoop1: TCP in base x=138.504 y=-514.48 z=214.154 mm, rx=-0.1348 ry=1.5599 rz=-0.0592 rad; joints [-39.422, -130.004, -76.262, -153.157, 47.788, -83.41] deg
                Waypoint ftr_scoop2: motionParameters(jointSpeed=1.047198 jointAcceleration=1.396263 cartesianSpeed=0.1 cartesianAcceleration=0.4); TCP in base x=194.287 y=-495.78 z=282.072 mm, rx=-0.179 ry=1.6121 rz=-0.016 rad; joints [-34.133, -129.723, -68.393, -165.549, 50.138, -80.843] deg
                Waypoint Waypoint_63: motionParameters(blendRadius=0.05); TCP in base x=101.295 y=-465.376 z=381.756 mm, rx=0.9726 ry=-0.1584 rz=2.8872 rad; joints [-48.863, -99.659, -71.872, -130.079, 68.56, 52.636] deg; TCP offset x=0 y=0 z=161 mm, rx=3.1415 ry=0 rz=0 rad
                Waypoint Start: motionParameters(jointSpeed=1.047198 jointAcceleration=1.396263 cartesianSpeed=0.15 cartesianAcceleration=0.6); TCP in base x=-33.065 y=-365.399 z=389.873 mm, rx=0 ry=0 rz=2.7258 rad; joints [-73.774, -70.638, -96.716, -102.629, 90.121, 40.001] deg; TCP offset x=0 y=0 z=161 mm, rx=3.1415 ry=0 rz=0 rad
                Popup Message (haltProgram=false message=Powder dispensed successfully... inputType=Text)
            SuppressedNode
              Script: tilt()
        SuppressedNode
          Script: tilt_send()
  '=========='
  Folder PostSettings [hidden by the author, left out]
